(* IEC 61131-3 sources: volt/packages/volt-lsp-iec/test-corpus/awa-palletizer/Device/Plc Logic/Application/Library Manager/CAA Behaviour Model, 13 files *)

(* ---- ERROR.dut ---- *)
TYPE ERROR :
(
	NO_ERROR,
	TIME_OUT
);
END_TYPE

(* ---- VERSIONCONSTANTS.gvl ---- *)
VAR_GLOBAL
	GC_BYVERSION : BYTE := 1;
	GC_BYVERSION_1 : BYTE := 0;
END_VAR

(* ---- IFBCOMMAND.itf ---- *)
INTERFACE IFBCOMMAND
END_INTERFACE

METHOD PRVABORT : BOOL
END_METHOD

METHOD PRVCYCLICACTION : BOOL
END_METHOD

METHOD PRVRESETOUTPUTS : BOOL
END_METHOD

METHOD PRVSTART : BOOL
END_METHOD

(* ---- GETSUPPLIERVERSION.pou ---- *)
FUNCTION GETSUPPLIERVERSION : WORD
VAR_INPUT
	XDUMMY : BOOL;
END_VAR
END_FUNCTION

(* ---- ETRIG.pou ---- *)
FUNCTION_BLOCK ETRIG
VAR_INPUT
	XEXECUTE : BOOL;
END_VAR
VAR_OUTPUT
	XDONE : BOOL;
	XBUSY : BOOL;
	XERROR : BOOL;
END_VAR
VAR
	XPREVIOUSEXECUTE : BOOL;
	XPREVIOUSABORTINPROGRESS : BOOL;
	XABORTINPROGRESS : BOOL;
	IERROR : INT;
END_VAR
END_FUNCTION_BLOCK

METHOD PRVABORT : BOOL
END_METHOD

METHOD PRVCYCLICACTION : BOOL
END_METHOD

METHOD PRVRESETOUTPUTS : BOOL
END_METHOD

METHOD PRVSTART : BOOL
END_METHOD

(* ---- ETRIGA.pou ---- *)
FUNCTION_BLOCK ETRIGA
VAR_INPUT
	XEXECUTE : BOOL;
	XABORT : BOOL;
END_VAR
VAR_OUTPUT
	XDONE : BOOL;
	XBUSY : BOOL;
	XERROR : BOOL;
	XABORTED : BOOL;
END_VAR
VAR
	XPREVIOUSABORTINPROGRESS : BOOL;
	XPREVIOUSEXECUTE : BOOL;
	XABORTINPROGRESS : BOOL;
	IERROR : INT;
END_VAR
END_FUNCTION_BLOCK

METHOD PRVABORT : BOOL
END_METHOD

METHOD PRVCYCLICACTION : BOOL
END_METHOD

METHOD PRVRESETOUTPUTS : BOOL
END_METHOD

METHOD PRVSTART : BOOL
END_METHOD

(* ---- ETRIGTL.pou ---- *)
FUNCTION_BLOCK ETRIGTL
VAR_INPUT
	XEXECUTE : BOOL;
	UDITIMELIMIT : UDINT;
END_VAR
VAR_OUTPUT
	XDONE : BOOL;
	XBUSY : BOOL;
	XERROR : BOOL;
END_VAR
VAR
	XPREVIOUSABORTINPROGRESS : BOOL;
	XPREVIOUSEXECUTE : BOOL;
	XABORTINPROGRESS : BOOL;
	XREPEAT : BOOL;
	TKFBSTART : CAA.TICK;
	TKTIMELIMIT : CAA.TICK;
	IERROR : INT;
END_VAR
END_FUNCTION_BLOCK

METHOD PRVABORT : BOOL
END_METHOD

METHOD PRVCYCLICACTION : BOOL
END_METHOD

METHOD PRVRESETOUTPUTS : BOOL
END_METHOD

METHOD PRVSTART : BOOL
END_METHOD

(* ---- ETRIGTLA.pou ---- *)
FUNCTION_BLOCK ETRIGTLA
VAR_INPUT
	XEXECUTE : BOOL;
	XABORT : BOOL;
	UDITIMELIMIT : UDINT;
END_VAR
VAR_OUTPUT
	XDONE : BOOL;
	XBUSY : BOOL;
	XERROR : BOOL;
	XABORTED : BOOL;
END_VAR
VAR
	XPREVIOUSABORTINPROGRESS : BOOL;
	XPREVIOUSEXECUTE : BOOL;
	XABORTINPROGRESS : BOOL;
	XREPEAT : BOOL;
	TKFBSTART : CAA.TICK;
	TKTIMELIMIT : CAA.TICK;
	IERROR : INT;
END_VAR
END_FUNCTION_BLOCK

METHOD PRVABORT : BOOL
END_METHOD

METHOD PRVCYCLICACTION : BOOL
END_METHOD

METHOD PRVRESETOUTPUTS : BOOL
END_METHOD

METHOD PRVSTART : BOOL
END_METHOD

(* ---- ETRIGTO.pou ---- *)
FUNCTION_BLOCK ETRIGTO
VAR_INPUT
	XEXECUTE : BOOL;
	UDITIMEOUT : UDINT;
END_VAR
VAR_OUTPUT
	XDONE : BOOL;
	XBUSY : BOOL;
	XERROR : BOOL;
END_VAR
VAR
	XPREVIOUSABORTINPROGRESS : BOOL;
	XPREVIOUSEXECUTE : BOOL;
	XABORTINPROGRESS : BOOL;
	TKSTART : CAA.TICK;
	TKTIMEOUT : CAA.TICK;
	IERROR : INT;
END_VAR
END_FUNCTION_BLOCK

METHOD PRVABORT : BOOL
END_METHOD

METHOD PRVCYCLICACTION : BOOL
END_METHOD

METHOD PRVRESETOUTPUTS : BOOL
END_METHOD

METHOD PRVSTART : BOOL
END_METHOD

(* ---- ETRIGTOA.pou ---- *)
FUNCTION_BLOCK ETRIGTOA
VAR_INPUT
	XEXECUTE : BOOL;
	XABORT : BOOL;
	UDITIMEOUT : UDINT;
END_VAR
VAR_OUTPUT
	XDONE : BOOL;
	XBUSY : BOOL;
	XERROR : BOOL;
	XABORTED : BOOL;
END_VAR
VAR
	XPREVIOUSABORTINPROGRESS : BOOL;
	XPREVIOUSEXECUTE : BOOL;
	XABORTINPROGRESS : BOOL;
	TKSTART : CAA.TICK;
	TKTIMEOUT : CAA.TICK;
	IERROR : INT;
END_VAR
END_FUNCTION_BLOCK

METHOD PRVABORT : BOOL
END_METHOD

METHOD PRVCYCLICACTION : BOOL
END_METHOD

METHOD PRVRESETOUTPUTS : BOOL
END_METHOD

METHOD PRVSTART : BOOL
END_METHOD

(* ---- ETRIGTOTL.pou ---- *)
FUNCTION_BLOCK ETRIGTOTL
VAR_INPUT
	XEXECUTE : BOOL;
	UDITIMELIMIT : UDINT;
	UDITIMEOUT : UDINT;
END_VAR
VAR_OUTPUT
	XDONE : BOOL;
	XBUSY : BOOL;
	XERROR : BOOL;
END_VAR
VAR
	XPREVIOUSABORTINPROGRESS : BOOL;
	XPREVIOUSEXECUTE : BOOL;
	XABORTINPROGRESS : BOOL;
	XREPEAT : BOOL;
	TKFBSTART : CAA.TICK;
	TKSTART : CAA.TICK;
	TKTIMELIMIT : CAA.TICK;
	TKTIMEOUT : CAA.TICK;
	IERROR : INT;
END_VAR
END_FUNCTION_BLOCK

METHOD PRVABORT : BOOL
END_METHOD

METHOD PRVCYCLICACTION : BOOL
END_METHOD

METHOD PRVRESETOUTPUTS : BOOL
END_METHOD

METHOD PRVSTART : BOOL
END_METHOD

(* ---- ETRIGTOTLA.pou ---- *)
FUNCTION_BLOCK ETRIGTOTLA
VAR_INPUT
	XEXECUTE : BOOL;
	XABORT : BOOL;
	UDITIMELIMIT : UDINT;
	UDITIMEOUT : UDINT;
END_VAR
VAR_OUTPUT
	XDONE : BOOL;
	XBUSY : BOOL;
	XERROR : BOOL;
	XABORTED : BOOL;
END_VAR
VAR
	XPREVIOUSABORTINPROGRESS : BOOL;
	XPREVIOUSEXECUTE : BOOL;
	XABORTINPROGRESS : BOOL;
	XREPEAT : BOOL;
	TKFBSTART : CAA.TICK;
	TKSTART : CAA.TICK;
	TKTIMELIMIT : CAA.TICK;
	TKTIMEOUT : CAA.TICK;
	IERROR : ERROR;
END_VAR
END_FUNCTION_BLOCK

METHOD PRVABORT : BOOL
END_METHOD

METHOD PRVCYCLICACTION : BOOL
END_METHOD

METHOD PRVRESETOUTPUTS : BOOL
END_METHOD

METHOD PRVSTART : BOOL
END_METHOD

(* ---- LTRIG.pou ---- *)
FUNCTION_BLOCK LTRIG
VAR_INPUT
	XENABLE : BOOL;
END_VAR
VAR_OUTPUT
	XDONE : BOOL;
	XBUSY : BOOL;
	XERROR : BOOL;
END_VAR
VAR
	XPREVIOUSABORTINPROGRESS : BOOL;
	XPREVIOUSENABLE : BOOL;
	XABORTINPROGRESS : BOOL;
	IERROR : INT;
END_VAR
END_FUNCTION_BLOCK

METHOD PRVABORT : BOOL
END_METHOD

METHOD PRVCYCLICACTION : BOOL
END_METHOD

METHOD PRVRESETOUTPUTS : BOOL
END_METHOD

METHOD PRVSTART : BOOL
END_METHOD
